   ElseIf Barcode = "D084" Then
       shell.Run "C:\Users\poh25\Videos\mini\D084.mp4"
   
   ElseIf Barcode = "D085" Then
       shell.Run "C:\Users\poh25\Videos\mini\D085.mp4"
   
   ElseIf Barcode = "D086" Then
       shell.Run "C:\Users\poh25\Videos\mini\D086.mp4"
   
   ElseIf Barcode = "D087" Then
       shell.Run "C:\Users\poh25\Videos\mini\D087.mp4"
   
   ElseIf Barcode = "D088" Then
       shell.Run "C:\Users\poh25\Videos\mini\D088.mp4"
   
   ElseIf Barcode = "D089" Then
       shell.Run "C:\Users\poh25\Videos\mini\D089.mp4"
   
   ElseIf Barcode = "D090" Then
       shell.Run "C:\Users\poh25\Videos\mini\D090.mp4"
   
   ElseIf Barcode = "D091" Then
       shell.Run "C:\Users\poh25\Videos\mini\D091.mp4"
   
   ElseIf Barcode = "D092" Then
       shell.Run "C:\Users\poh25\Videos\mini\D092.mp4"
   
   ElseIf Barcode = "D093" Then
       shell.Run "C:\Users\poh25\Videos\mini\D093.mp4"
   
   ElseIf Barcode = "D094" Then
       shell.Run "C:\Users\poh25\Videos\mini\D094.mp4"
   
   ElseIf Barcode = "D095" Then
       shell.Run "C:\Users\poh25\Videos\mini\D095.mp4"
   
   ElseIf Barcode = "D096" Then
       shell.Run "C:\Users\poh25\Videos\mini\D096.mp4"
   
   ElseIf Barcode = "D097" Then
       shell.Run "C:\Users\poh25\Videos\mini\D097.mp4"
   
   ElseIf Barcode = "D098" Then
       shell.Run "C:\Users\poh25\Videos\mini\D098.mp4"
   
   ElseIf Barcode = "D099" Then
       shell.Run "C:\Users\poh25\Videos\mini\D099.mp4"
   
   ElseIf Barcode = "D100" Then
       shell.Run "C:\Users\poh25\Videos\mini\D100.mp4"
   
   ElseIf Barcode = "E001" Then
       shell.Run "C:\Users\poh25\Videos\mini\E001.mp4"
   
   ElseIf Barcode = "E002" Then
       shell.Run "C:\Users\poh25\Videos\mini\E002.mp4"
   
   ElseIf Barcode = "E003" Then
       shell.Run "C:\Users\poh25\Videos\mini\E003.mp4"
   
   ElseIf Barcode = "E004" Then
       shell.Run "C:\Users\poh25\Videos\mini\E004.mp4"
   
   ElseIf Barcode = "E005" Then
       shell.Run "C:\Users\poh25\Videos\mini\E005.mp4"
   
   ElseIf Barcode = "E006" Then
       shell.Run "C:\Users\poh25\Videos\mini\E006.mp4"
   
   ElseIf Barcode = "E007" Then
       shell.Run "C:\Users\poh25\Videos\mini\E007.mp4"
   
   ElseIf Barcode = "E008" Then
       shell.Run "C:\Users\poh25\Videos\mini\E008.mp4"
   
   ElseIf Barcode = "E009" Then
       shell.Run "C:\Users\poh25\Videos\mini\E009.mp4"
   
   ElseIf Barcode = "E010" Then
       shell.Run "C:\Users\poh25\Videos\mini\E010.mp4"
   
   ElseIf Barcode = "E011" Then
       shell.Run "C:\Users\poh25\Videos\mini\E011.mp4"
   
   ElseIf Barcode = "E012" Then
       shell.Run "C:\Users\poh25\Videos\mini\E012.mp4"
   
   ElseIf Barcode = "E013" Then
       shell.Run "C:\Users\poh25\Videos\mini\E013.mp4"
   
   ElseIf Barcode = "E014" Then
       shell.Run "C:\Users\poh25\Videos\mini\E014.mp4"
   
   ElseIf Barcode = "E015" Then
       shell.Run "C:\Users\poh25\Videos\mini\E015.mp4"
   
   ElseIf Barcode = "E016" Then
       shell.Run "C:\Users\poh25\Videos\mini\E016.mp4"
   
   ElseIf Barcode = "E017" Then
       shell.Run "C:\Users\poh25\Videos\mini\E017.mp4"
   
   ElseIf Barcode = "E018" Then
       shell.Run "C:\Users\poh25\Videos\mini\E018.mp4"
   
   ElseIf Barcode = "E019" Then
       shell.Run "C:\Users\poh25\Videos\mini\E019.mp4"
   
   ElseIf Barcode = "E020" Then
       shell.Run "C:\Users\poh25\Videos\mini\E020.mp4"
   
   ElseIf Barcode = "E021" Then
       shell.Run "C:\Users\poh25\Videos\mini\E021.mp4"
   
   ElseIf Barcode = "E022" Then
       shell.Run "C:\Users\poh25\Videos\mini\E022.mp4"
   
   ElseIf Barcode = "E023" Then
       shell.Run "C:\Users\poh25\Videos\mini\E023.mp4"
   
   ElseIf Barcode = "E024" Then
       shell.Run "C:\Users\poh25\Videos\mini\E024.mp4"
   
   ElseIf Barcode = "E025" Then
       shell.Run "C:\Users\poh25\Videos\mini\E025.mp4"
   
   ElseIf Barcode = "E026" Then
       shell.Run "C:\Users\poh25\Videos\mini\E026.mp4"
   
   ElseIf Barcode = "E027" Then
       shell.Run "C:\Users\poh25\Videos\mini\E027.mp4"
   
   ElseIf Barcode = "E028" Then
       shell.Run "C:\Users\poh25\Videos\mini\E028.mp4"
   
   ElseIf Barcode = "E029" Then
       shell.Run "C:\Users\poh25\Videos\mini\E029.mp4"
   
   ElseIf Barcode = "E030" Then
       shell.Run "C:\Users\poh25\Videos\mini\E030.mp4"
   
   ElseIf Barcode = "E031" Then
       shell.Run "C:\Users\poh25\Videos\mini\E031.mp4"
   
   ElseIf Barcode = "E032" Then
       shell.Run "C:\Users\poh25\Videos\mini\E032.mp4"
   
   ElseIf Barcode = "E033" Then
       shell.Run "C:\Users\poh25\Videos\mini\E033.mp4"
   
   ElseIf Barcode = "E034" Then
       shell.Run "C:\Users\poh25\Videos\mini\E034.mp4"
   
   ElseIf Barcode = "E035" Then
       shell.Run "C:\Users\poh25\Videos\mini\E035.mp4"
   
   ElseIf Barcode = "E036" Then
       shell.Run "C:\Users\poh25\Videos\mini\E036.mp4"
   
   ElseIf Barcode = "E037" Then
       shell.Run "C:\Users\poh25\Videos\mini\E037.mp4"
   
   ElseIf Barcode = "E038" Then
       shell.Run "C:\Users\poh25\Videos\mini\E038.mp4"
   
   ElseIf Barcode = "E039" Then
       shell.Run "C:\Users\poh25\Videos\mini\E039.mp4"
   
   ElseIf Barcode = "E040" Then
       shell.Run "C:\Users\poh25\Videos\mini\E040.mp4"
   
   ElseIf Barcode = "E041" Then
       shell.Run "C:\Users\poh25\Videos\mini\E041.mp4"
   
   ElseIf Barcode = "E042" Then
       shell.Run "C:\Users\poh25\Videos\mini\E042.mp4"
   
   ElseIf Barcode = "E043" Then
       shell.Run "C:\Users\poh25\Videos\mini\E043.mp4"
   
   ElseIf Barcode = "E044" Then
       shell.Run "C:\Users\poh25\Videos\mini\E044.mp4"
   
   ElseIf Barcode = "E045" Then
       shell.Run "C:\Users\poh25\Videos\mini\E045.mp4"
   
   ElseIf Barcode = "E046" Then
       shell.Run "C:\Users\poh25\Videos\mini\E046.mp4"
   
   ElseIf Barcode = "E047" Then
       shell.Run "C:\Users\poh25\Videos\mini\E047.mp4"
   
   ElseIf Barcode = "E048" Then
       shell.Run "C:\Users\poh25\Videos\mini\E048.mp4"
   
   ElseIf Barcode = "E049" Then
       shell.Run "C:\Users\poh25\Videos\mini\E049.mp4"
   
   ElseIf Barcode = "E050" Then
       shell.Run "C:\Users\poh25\Videos\mini\E050.mp4"
   
   ElseIf Barcode = "E051" Then
       shell.Run "C:\Users\poh25\Videos\mini\E051.mp4"
   
   ElseIf Barcode = "E052" Then
       shell.Run "C:\Users\poh25\Videos\mini\E052.mp4"
   
   ElseIf Barcode = "E053" Then
       shell.Run "C:\Users\poh25\Videos\mini\E053.mp4"
   
   ElseIf Barcode = "E054" Then
       shell.Run "C:\Users\poh25\Videos\mini\E054.mp4"
   
   ElseIf Barcode = "E055" Then
       shell.Run "C:\Users\poh25\Videos\mini\E055.mp4"
   
   ElseIf Barcode = "E056" Then
       shell.Run "C:\Users\poh25\Videos\mini\E056.mp4"
   
   ElseIf Barcode = "E057" Then
       shell.Run "C:\Users\poh25\Videos\mini\E057.mp4"
   
   ElseIf Barcode = "E058" Then
       shell.Run "C:\Users\poh25\Videos\mini\E058.mp4"
   
   ElseIf Barcode = "E059" Then
       shell.Run "C:\Users\poh25\Videos\mini\E059.mp4"
   
   ElseIf Barcode = "E060" Then
       shell.Run "C:\Users\poh25\Videos\mini\E060.mp4"
   
   ElseIf Barcode = "E061" Then
       shell.Run "C:\Users\poh25\Videos\mini\E061.mp4"
   
   ElseIf Barcode = "E062" Then
       shell.Run "C:\Users\poh25\Videos\mini\E062.mp4"
   
   ElseIf Barcode = "E063" Then
       shell.Run "C:\Users\poh25\Videos\mini\E063.mp4"
   
   ElseIf Barcode = "E064" Then
       shell.Run "C:\Users\poh25\Videos\mini\E064.mp4"
   
   ElseIf Barcode = "E065" Then
       shell.Run "C:\Users\poh25\Videos\mini\E065.mp4"
   
   ElseIf Barcode = "E066" Then
       shell.Run "C:\Users\poh25\Videos\mini\E066.mp4"
   
   ElseIf Barcode = "E067" Then
       shell.Run "C:\Users\poh25\Videos\mini\E067.mp4"
   
   ElseIf Barcode = "E068" Then
       shell.Run "C:\Users\poh25\Videos\mini\E068.mp4"
   
   ElseIf Barcode = "E069" Then
       shell.Run "C:\Users\poh25\Videos\mini\E069.mp4"
   
   ElseIf Barcode = "E070" Then
       shell.Run "C:\Users\poh25\Videos\mini\E070.mp4"
   
   ElseIf Barcode = "E071" Then
       shell.Run "C:\Users\poh25\Videos\mini\E071.mp4"
   
   ElseIf Barcode = "E072" Then
       shell.Run "C:\Users\poh25\Videos\mini\E072.mp4"
   
   ElseIf Barcode = "E073" Then
       shell.Run "C:\Users\poh25\Videos\mini\E073.mp4"
   
   ElseIf Barcode = "E074" Then
       shell.Run "C:\Users\poh25\Videos\mini\E074.mp4"
   
   ElseIf Barcode = "E075" Then
       shell.Run "C:\Users\poh25\Videos\mini\E075.mp4"
   
   ElseIf Barcode = "E076" Then
       shell.Run "C:\Users\poh25\Videos\mini\E076.mp4"
   
   ElseIf Barcode = "E077" Then
       shell.Run "C:\Users\poh25\Videos\mini\E077.mp4"
   
   ElseIf Barcode = "E078" Then
       shell.Run "C:\Users\poh25\Videos\mini\E078.mp4"
   
   ElseIf Barcode = "E079" Then
       shell.Run "C:\Users\poh25\Videos\mini\E079.mp4"
   
   ElseIf Barcode = "E080" Then
       shell.Run "C:\Users\poh25\Videos\mini\E080.mp4"
   
   ElseIf Barcode = "E081" Then
       shell.Run "C:\Users\poh25\Videos\mini\E081.mp4"
   
   ElseIf Barcode = "E082" Then
       shell.Run "C:\Users\poh25\Videos\mini\E082.mp4"
   
   ElseIf Barcode = "E083" Then
       shell.Run "C:\Users\poh25\Videos\mini\E083.mp4"
   
   ElseIf Barcode = "E084" Then
       shell.Run "C:\Users\poh25\Videos\mini\E084.mp4"
   
   ElseIf Barcode = "E085" Then
       shell.Run "C:\Users\poh25\Videos\mini\E085.mp4"
   
   ElseIf Barcode = "E086" Then
       shell.Run "C:\Users\poh25\Videos\mini\E086.mp4"
   
   ElseIf Barcode = "E087" Then
       shell.Run "C:\Users\poh25\Videos\mini\E087.mp4"
   
   ElseIf Barcode = "E088" Then
       shell.Run "C:\Users\poh25\Videos\mini\E088.mp4"
   
   ElseIf Barcode = "E089" Then
       shell.Run "C:\Users\poh25\Videos\mini\E089.mp4"
   
   ElseIf Barcode = "E090" Then
       shell.Run "C:\Users\poh25\Videos\mini\E090.mp4"
   
   ElseIf Barcode = "E091" Then
       shell.Run "C:\Users\poh25\Videos\mini\E091.mp4"
   
   ElseIf Barcode = "E092" Then
       shell.Run "C:\Users\poh25\Videos\mini\E092.mp4"
   
   ElseIf Barcode = "E093" Then
       shell.Run "C:\Users\poh25\Videos\mini\E093.mp4"
   
   ElseIf Barcode = "E094" Then
       shell.Run "C:\Users\poh25\Videos\mini\E094.mp4"
   
   ElseIf Barcode = "E095" Then
       shell.Run "C:\Users\poh25\Videos\mini\E095.mp4"
   
   ElseIf Barcode = "E096" Then
       shell.Run "C:\Users\poh25\Videos\mini\E096.mp4"
   
   ElseIf Barcode = "E097" Then
       shell.Run "C:\Users\poh25\Videos\mini\E097.mp4"
   
   ElseIf Barcode = "E098" Then
       shell.Run "C:\Users\poh25\Videos\mini\E098.mp4"
   
   ElseIf Barcode = "E099" Then
       shell.Run "C:\Users\poh25\Videos\mini\E099.mp4"
   
   ElseIf Barcode = "E100" Then
       shell.Run "C:\Users\poh25\Videos\mini\E100.mp4"
   
   ElseIf Barcode = "F001" Then
       shell.Run "C:\Users\poh25\Videos\mini\F001.mp4"
   
   ElseIf Barcode = "F002" Then
       shell.Run "C:\Users\poh25\Videos\mini\F002.mp4"
   
   ElseIf Barcode = "F003" Then
       shell.Run "C:\Users\poh25\Videos\mini\F003.mp4"
   
   ElseIf Barcode = "F004" Then
       shell.Run "C:\Users\poh25\Videos\mini\F004.mp4"
   
   ElseIf Barcode = "F005" Then
       shell.Run "C:\Users\poh25\Videos\mini\F005.mp4"
   
   ElseIf Barcode = "F006" Then
       shell.Run "C:\Users\poh25\Videos\mini\F006.mp4"
   
   ElseIf Barcode = "F007" Then
       shell.Run "C:\Users\poh25\Videos\mini\F007.mp4"
   
   ElseIf Barcode = "F008" Then
       shell.Run "C:\Users\poh25\Videos\mini\F008.mp4"
   
   ElseIf Barcode = "F009" Then
       shell.Run "C:\Users\poh25\Videos\mini\F009.mp4"
   
   ElseIf Barcode = "F010" Then
       shell.Run "C:\Users\poh25\Videos\mini\F010.mp4"
   
   ElseIf Barcode = "F011" Then
       shell.Run "C:\Users\poh25\Videos\mini\F011.mp4"
   
   ElseIf Barcode = "F012" Then
       shell.Run "C:\Users\poh25\Videos\mini\F012.mp4"
   
   ElseIf Barcode = "F013" Then
       shell.Run "C:\Users\poh25\Videos\mini\F013.mp4"
   
   ElseIf Barcode = "F014" Then
       shell.Run "C:\Users\poh25\Videos\mini\F014.mp4"
   
   ElseIf Barcode = "F015" Then
       shell.Run "C:\Users\poh25\Videos\mini\F015.mp4"
   
   ElseIf Barcode = "F016" Then
       shell.Run "C:\Users\poh25\Videos\mini\F016.mp4"
   
   ElseIf Barcode = "F017" Then
       shell.Run "C:\Users\poh25\Videos\mini\F017.mp4"
   
   ElseIf Barcode = "F018" Then
       shell.Run "C:\Users\poh25\Videos\mini\F018.mp4"
   
   ElseIf Barcode = "F019" Then
       shell.Run "C:\Users\poh25\Videos\mini\F019.mp4"
   
   ElseIf Barcode = "F020" Then
       shell.Run "C:\Users\poh25\Videos\mini\F020.mp4"
   
   End If
   
   Set shell = Nothing
*)